DATA_BLOCK "FRK_AccessPolicies"
{ S7_Optimized_Access := 'TRUE' }
VERSION : 0.1
NON_RETAIN
VAR RETAIN
    Rows {ExternalAccessible := 'False'; ExternalVisible := 'False'; ExternalWritable := 'False'} : Array[1..1] of "FRK_AccessPolicyImage";
END_VAR
BEGIN
END_DATA_BLOCK
